(* IEC 61131-3 sources: canworks/examples/virtual-plant/pous/programs, 3 files *)

(* ---- canworks_in.st ---- *)
PROGRAM canworks_in
  VAR
    i0  : WORD AT %IW100; (* cw_map_hash *)
    i1  : WORD AT %IW101; (* cw_map_hash_w1 *)
    i2  : WORD AT %IW102; (* cw_status *)
    i3  : WORD AT %IW103; (* cw_status_w1 *)
    i4  : WORD AT %IW104; (* cw_status_w2 *)
    i5  : WORD AT %IW105; (* cw_status_w3 *)
    i6  : WORD AT %IW106; (* io_rtd_AI0_Input_PV *)
    i7  : WORD AT %IW107; (* io_rtd_AI1_Input_PV *)
    i8  : WORD AT %IW108; (* io_rtd_AI2_Input_PV *)
    i9  : WORD AT %IW109; (* io_rtd_AI3_Input_PV *)
    i10 : WORD AT %IW110; (* io_dio_Read_input_8_bit_1 *)
    i11 : WORD AT %IW111; (* io_dio_Read_analogue_input_1 *)
    i12 : WORD AT %IW112; (* io_dio_Read_analogue_input_2 *)
    i13 : WORD AT %IW113; (* io_dio_operating_hours *)
    i14 : WORD AT %IW114; (* io_dio_operating_hours_w1 *)
    i15 : WORD AT %IW115; (* io_new_io_Read_input_8_bit_1 *)
    i16 : WORD AT %IW116; (* motion_conveyor_speed_actual *)
    i17 : WORD AT %IW117; (* motion_conveyor_belt_position *)
    i18 : WORD AT %IW118; (* motion_conveyor_belt_position_w1 *)
    i19 : WORD AT %IW119; (* host_cell_alarm *)
    i20 : WORD AT %IW120; (* cell_temp_limit *)
    i21 : WORD AT %IW121; (* host_cell_belt_position *)
    i22 : WORD AT %IW122; (* host_cell_belt_position_w1 *)
    i23 : WORD AT %IW123; (* host_cell_cycle_count *)
    i24 : WORD AT %IW124; (* host_cell_cycle_count_w1 *)
    i25 : WORD AT %IW125; (* host_cell_temperature *)
    i26 : WORD AT %IW126; (* host_cell_Nodes_0_31 *)
    i27 : WORD AT %IW127; (* host_cell_Nodes_0_31_w1 *)
    i28 : WORD AT %IW128; (* host_cell_Nodes_0_31_2 *)
    i29 : WORD AT %IW129; (* host_cell_Nodes_0_31_2_w1 *)
    i30 : WORD AT %IW130; (* io_can_bus_state *)
    i31 : WORD AT %IW131; (* io_rtd_ok *)
    i32 : WORD AT %IW132; (* io_rtd_emcy *)
    i33 : WORD AT %IW133; (* io_dio_state *)
    i34 : WORD AT %IW134; (* io_dio_emcy *)
    i35 : WORD AT %IW135; (* io_dio_operating_hours_status *)
    i36 : WORD AT %IW136; (* motion_can_master_state *)
    i37 : WORD AT %IW137; (* motion_conveyor_emcy *)
    i38 : WORD AT %IW138; (* host_can_master_state *)
    i39 : WORD AT %IW139; (* host_cell_state *)
    i40 : WORD AT %IW140; (* host_cell_emcy *)
    i41 : WORD AT %IW141; (* cw_live_list_io *)
    i42 : WORD AT %IW142; (* cw_live_list_io_w1 *)
    i43 : WORD AT %IW143; (* cw_live_list_io_w2 *)
    i44 : WORD AT %IW144; (* cw_live_list_io_w3 *)
    i45 : WORD AT %IW145; (* cw_live_list_io_w4 *)
    i46 : WORD AT %IW146; (* cw_live_list_io_w5 *)
    i47 : WORD AT %IW147; (* cw_live_list_io_w6 *)
    i48 : WORD AT %IW148; (* cw_live_list_io_w7 *)
    i49 : WORD AT %IW149; (* cw_live_list_motion *)
    i50 : WORD AT %IW150; (* cw_live_list_motion_w1 *)
    i51 : WORD AT %IW151; (* cw_live_list_motion_w2 *)
    i52 : WORD AT %IW152; (* cw_live_list_motion_w3 *)
    i53 : WORD AT %IW153; (* cw_live_list_motion_w4 *)
    i54 : WORD AT %IW154; (* cw_live_list_motion_w5 *)
    i55 : WORD AT %IW155; (* cw_live_list_motion_w6 *)
    i56 : WORD AT %IW156; (* cw_live_list_motion_w7 *)
    i57 : WORD AT %IW157; (* cw_live_list_host *)
    i58 : WORD AT %IW158; (* cw_live_list_host_w1 *)
    i59 : WORD AT %IW159; (* cw_live_list_host_w2 *)
    i60 : WORD AT %IW160; (* cw_live_list_host_w3 *)
    i61 : WORD AT %IW161; (* cw_live_list_host_w4 *)
    i62 : WORD AT %IW162; (* cw_live_list_host_w5 *)
    i63 : WORD AT %IW163; (* cw_live_list_host_w6 *)
    i64 : WORD AT %IW164; (* cw_live_list_host_w7 *)
    i65 : WORD AT %IW165; (* cw_sdo_bridge_response *)
    i66 : WORD AT %IW166; (* cw_sdo_bridge_response_w1 *)
    i67 : WORD AT %IW167; (* cw_sdo_bridge_response_w2 *)
    i68 : WORD AT %IW168; (* cw_sdo_bridge_response_w3 *)
    i69 : WORD AT %IW169; (* cw_sdo_bridge_response_w4 *)
    i70 : WORD AT %IW170; (* cw_sdo_bridge_response_w5 *)
    i71 : WORD AT %IW171; (* cw_sdo_bridge_response_w6 *)
  END_VAR
  VAR
    last_counter : WORD;
    moved        : BOOL;
    stale        : TON;
  END_VAR

(* Generated by canworks from canworks/canworks.json: do not edit, Save rewrites it. *)
moved := i3 <> last_counter;
last_counter := i3;
stale(IN := NOT moved, PT := T#300ms);
canworks.ok := i0 = WORD#16#662D AND i1 = WORD#16#449C AND NOT stale.Q;
canworks.bus_ok := canworks.ok AND (i5 AND WORD#16#0002) = WORD#0;
canworks.link[21] := WORD#16#0B06 OR SEL(canworks.ok, WORD#0, WORD#1);
canworks.link[0] := i2;
canworks.link[1] := i3;
canworks.link[2] := i4;
canworks.link[3] := i5;
canworks.link[14] := i65;
canworks.link[15] := i66;
canworks.link[16] := i67;
canworks.link[17] := i68;
canworks.link[18] := i69;
canworks.link[19] := i70;
canworks.link[20] := i71;
canworks.link[25] := i41;
canworks.link[26] := i42;
canworks.link[27] := i43;
canworks.link[28] := i44;
canworks.link[29] := i45;
canworks.link[30] := i46;
canworks.link[31] := i47;
canworks.link[32] := i48;
canworks.link[33] := i49;
canworks.link[34] := i50;
canworks.link[35] := i51;
canworks.link[36] := i52;
canworks.link[37] := i53;
canworks.link[38] := i54;
canworks.link[39] := i55;
canworks.link[40] := i56;
canworks.link[49] := i57;
canworks.link[50] := i58;
canworks.link[51] := i59;
canworks.link[52] := i60;
canworks.link[53] := i61;
canworks.link[54] := i62;
canworks.link[55] := i63;
canworks.link[56] := i64;
canworks.io_can_bus_state := SEL(canworks.ok, USINT#0, WORD_TO_USINT((i30 AND WORD#16#00FF)));
canworks.io_can_master_state := SEL(canworks.ok, USINT#0, WORD_TO_USINT(SHR(i30, 8)));
canworks.motion_can_master_state := SEL(canworks.ok, USINT#0, WORD_TO_USINT(SHR(i36, 8)));
canworks.host_can_master_state := SEL(canworks.ok, USINT#0, WORD_TO_USINT((i38 AND WORD#16#00FF)));
canworks.io_rtd_ok := SEL(canworks.ok, FALSE, (i31 AND WORD#16#0100) <> WORD#0);
canworks.io_rtd_state := SEL(canworks.ok, USINT#0, WORD_TO_USINT((i31 AND WORD#16#00FF)));
canworks.io_rtd_emcy := SEL(canworks.ok, WORD#0, i32);
canworks.io_rtd_tpdo1_timeout := SEL(canworks.ok, FALSE, (i31 AND WORD#16#0200) <> WORD#0);
canworks.io_rtd_AI0_Input_PV := WORD_TO_INT(i6);
canworks.io_rtd_AI1_Input_PV := WORD_TO_INT(i7);
canworks.io_rtd_AI2_Input_PV := WORD_TO_INT(i8);
canworks.io_rtd_AI3_Input_PV := WORD_TO_INT(i9);
canworks.io_dio_ok := SEL(canworks.ok, FALSE, (i31 AND WORD#16#0400) <> WORD#0);
canworks.io_dio_state := SEL(canworks.ok, USINT#0, WORD_TO_USINT(SHR(i33, 8)));
canworks.io_dio_emcy := SEL(canworks.ok, WORD#0, i34);
canworks.io_dio_Read_input_8_bit_1 := WORD_TO_USINT(SHR(i10, 8));
canworks.io_dio_Read_input_8_bit_2 := WORD_TO_USINT((i10 AND WORD#16#00FF));
canworks.io_dio_Read_analogue_input_1 := WORD_TO_INT(i11);
canworks.io_dio_Read_analogue_input_2 := WORD_TO_INT(i12);
canworks.io_dio_operating_hours := DWORD_TO_UDINT((SHL(WORD_TO_DWORD(i14), 16) OR WORD_TO_DWORD(i13)));
canworks.io_dio_operating_hours_status := SEL(canworks.ok, USINT#0, WORD_TO_USINT(SHR(i35, 8)));
canworks.io_dio_filter_time_status := SEL(canworks.ok, USINT#0, WORD_TO_USINT((i35 AND WORD#16#00FF)));
canworks.io_new_io_ok := SEL(canworks.ok, FALSE, (i31 AND WORD#16#0800) <> WORD#0);
canworks.io_new_io_Read_input_8_bit_1 := WORD_TO_USINT(SHR(i15, 8));
canworks.motion_conveyor_ok := SEL(canworks.ok, FALSE, (i31 AND WORD#16#1000) <> WORD#0);
canworks.motion_conveyor_state := SEL(canworks.ok, USINT#0, WORD_TO_USINT((i36 AND WORD#16#00FF)));
canworks.motion_conveyor_emcy := SEL(canworks.ok, WORD#0, i37);
canworks.motion_conveyor_speed_actual := WORD_TO_INT(i16);
canworks.motion_conveyor_belt_position := DWORD_TO_DINT((SHL(WORD_TO_DWORD(i18), 16) OR WORD_TO_DWORD(i17)));
canworks.host_cell_ok := SEL(canworks.ok, FALSE, (i31 AND WORD#16#4000) <> WORD#0);
canworks.host_cell_state := SEL(canworks.ok, USINT#0, WORD_TO_USINT(SHR(i39, 8)));
canworks.host_cell_emcy := SEL(canworks.ok, WORD#0, i40);
canworks.host_cell_alarm := (i19 AND WORD#16#0200) <> WORD#0;
canworks.host_cell_belt_position := DWORD_TO_DINT((SHL(WORD_TO_DWORD(i22), 16) OR WORD_TO_DWORD(i21)));
canworks.host_cell_cycle_count := DWORD_TO_UDINT((SHL(WORD_TO_DWORD(i24), 16) OR WORD_TO_DWORD(i23)));
canworks.host_cell_temperature := WORD_TO_INT(i25);
canworks.host_cell_Nodes_0_31 := DWORD_TO_UDINT((SHL(WORD_TO_DWORD(i27), 16) OR WORD_TO_DWORD(i26)));
canworks.host_cell_Nodes_0_31_2 := DWORD_TO_UDINT((SHL(WORD_TO_DWORD(i29), 16) OR WORD_TO_DWORD(i28)));
canworks.cell_line_run := (i19 AND WORD#16#0100) <> WORD#0;
canworks.cell_temp_limit := WORD_TO_INT(i20);
canworks.cell_state := SEL(canworks.ok, USINT#0, WORD_TO_USINT(SHR(i38, 8)));
canworks.cell_comm_ok := SEL(canworks.ok, FALSE, (i31 AND WORD#16#2000) <> WORD#0);

END_PROGRAM

(* ---- canworks_out.st ---- *)
PROGRAM canworks_out
  VAR
    q0  : WORD AT %QW100; (* cw_plc_link *)
    q1  : WORD AT %QW101; (* cw_plc_link_w1 *)
    q2  : WORD AT %QW102; (* cw_plc_link_w2 *)
    q3  : WORD AT %QW103; (* io_dio_Write_output_8_bit_1 *)
    q4  : WORD AT %QW104; (* io_dio_Write_analogue_output_2 *)
    q5  : WORD AT %QW105; (* io_dio_filter_time *)
    q6  : WORD AT %QW106; (* io_new_io_Write_output_8_bit_1 *)
    q7  : WORD AT %QW107; (* motion_conveyor_speed_setpoint *)
    q8  : WORD AT %QW108; (* host_cell_line_run *)
    q9  : WORD AT %QW109; (* cell_belt_position *)
    q10 : WORD AT %QW110; (* cell_belt_position_w1 *)
    q11 : WORD AT %QW111; (* cell_cycle_count *)
    q12 : WORD AT %QW112; (* cell_cycle_count_w1 *)
    q13 : WORD AT %QW113; (* host_cell_temp_limit *)
    q14 : WORD AT %QW114; (* host_cell_analog_out *)
    q15 : WORD AT %QW115; (* io_dio_filter_time_trig *)
    q16 : WORD AT %QW116; (* cell_emcy *)
    q17 : WORD AT %QW117; (* cell_errreg *)
    q18 : WORD AT %QW118; (* cw_control *)
    q19 : WORD AT %QW119; (* cw_control_w1 *)
    q20 : WORD AT %QW120; (* cw_control_w2 *)
    q21 : WORD AT %QW121; (* cw_sdo_bridge_request *)
    q22 : WORD AT %QW122; (* cw_sdo_bridge_request_w1 *)
    q23 : WORD AT %QW123; (* cw_sdo_bridge_request_w2 *)
    q24 : WORD AT %QW124; (* cw_sdo_bridge_request_w3 *)
    q25 : WORD AT %QW125; (* cw_sdo_bridge_request_w4 *)
    q26 : WORD AT %QW126; (* cw_sdo_bridge_request_w5 *)
    q27 : WORD AT %QW127; (* cw_sdo_bridge_request_w6 *)
  END_VAR
  VAR
    d9  : DWORD;
    d11 : DWORD;
  END_VAR

(* Generated by canworks from canworks/canworks.json: do not edit, Save rewrites it. *)
d9 := DINT_TO_DWORD(canworks.cell_belt_position);
d11 := UDINT_TO_DWORD(canworks.cell_cycle_count);
q3 := SHL((USINT_TO_WORD(canworks.io_dio_Write_output_8_bit_1) AND WORD#16#00FF), 8) OR (USINT_TO_WORD(canworks.io_dio_Write_output_8_bit_2) AND WORD#16#00FF);
q4 := INT_TO_WORD(canworks.io_dio_Write_analogue_output_2);
q5 := UINT_TO_WORD(canworks.io_dio_filter_time);
q6 := SHL((USINT_TO_WORD(canworks.io_new_io_Write_output_8_bit_1) AND WORD#16#00FF), 8);
q7 := INT_TO_WORD(canworks.motion_conveyor_speed_setpoint);
q8 := SEL(canworks.host_cell_line_run, WORD#0, WORD#16#0200) OR SEL(canworks.cell_alarm, WORD#0, WORD#16#0100);
q9 := DWORD_TO_WORD(d9);
q10 := DWORD_TO_WORD(SHR(d9, 16));
q11 := DWORD_TO_WORD(d11);
q12 := DWORD_TO_WORD(SHR(d11, 16));
q13 := INT_TO_WORD(canworks.host_cell_temp_limit);
q14 := INT_TO_WORD(canworks.host_cell_analog_out);
q15 := SEL(canworks.io_dio_filter_time_trig, WORD#0, WORD#16#0100);
q16 := canworks.cell_emcy;
q17 := SHL((BYTE_TO_WORD(canworks.cell_errreg) AND WORD#16#00FF), 8);
q18 := canworks.link[4];
q19 := canworks.link[5];
q20 := canworks.link[6];
q21 := canworks.link[7];
q22 := canworks.link[8];
q23 := canworks.link[9];
q24 := canworks.link[10];
q25 := canworks.link[11];
q26 := canworks.link[12];
q27 := canworks.link[13];
(* PLC link header, last: running, then the map hash 0x662d449c *)
q1 := WORD#16#662D;
q2 := WORD#16#449C;
q0 := WORD#1;

END_PROGRAM

(* ---- main.st ---- *)
PROGRAM main
  VAR
    (* The demo (docs/tour.md). The CANopen values are in the `canworks`
       variable list, which canworks_in fills from the bridge before main and
       canworks_out sends after it (the configurator writes all three). *)
    temp_c          : REAL;   (* RTD channel 0 in degC (the module sends 0.1 degC) *)
    limit           : INT;    (* alarm limit in 0.1 degC, from the cell's upper master *)
    alarm           : BOOL;   (* channel 0 above the limit: DIO-16 output 0.0 and the cell's alarm *)
    fault           : BOOL;   (* a node lost, a PDO timed out or an EMCY active: new_io output 0.0 *)
    pattern         : USINT := 1;  (* running light on DIO-16 output byte 2, read back on input byte 2 *)
    tick            : INT;
    loop_errors     : UDINT;  (* times the read-back input did not follow the output *)
    loop_ok         : BOOL;
    cycles          : UDINT;
    restart_dio     : BOOL;   (* set it in the debugger: NMT reset of node dio (6) *)
    started         : BOOL;
    rd_product      : CO_SDO_READ;   (* network io (0), node 5: 0x1018:2 product code *)
    rd_conveyor     : CO_SDO_READ;   (* network motion (1), node 4: 0x1018:2 product code *)
    wr_ai_interrupt : CO_SDO_WRITE;  (* network io (0), node 6: 0x6423 analogue input global interrupt enable *)
    reset_dio       : CO_NMT;        (* network io (0), node 6: RESET NODE when restart_dio is set *)
    rtd_product     : UDINT;
    conveyor_product : UDINT;
    sdo_errors      : INT;
    (* The host network plays the cell's machine controller (the upper master). *)
    host_field_ok   : BOOL;   (* the gateway reports io nodes 5, 6, 7 and motion node 4 operational *)
    speed           : INT := 1000;  (* conveyor speed while the upper master runs the line *)
  END_VAR

(* Temperature, alarm and the I/O loopback on network io *)
cycles := cycles + 1;
canworks.cell_cycle_count := cycles;
temp_c := INT_TO_REAL(canworks.io_rtd_AI0_Input_PV) / 10.0;
limit := canworks.cell_temp_limit;
IF limit = 0 THEN limit := 250; END_IF  (* no upper master: 25.0 degC *)
alarm := canworks.io_rtd_ok AND canworks.io_rtd_AI0_Input_PV > limit;
canworks.cell_alarm := alarm;
IF alarm THEN
  canworks.cell_emcy := 16#4210;  (* temperature too high: the cell slave sends it once *)
  canworks.cell_errreg := 16#09;  (* generic + temperature *)
ELSE
  canworks.cell_emcy := 0;
  canworks.cell_errreg := 0;
END_IF
canworks.io_dio_Write_output_8_bit_1 := BOOL_TO_USINT(alarm);

(* DIO-16 loops its outputs back to its inputs: a running light on byte 2,
   checked a few PDO round trips later. *)
tick := tick + 1;
IF tick >= 25 THEN
  tick := 0;
  IF canworks.io_dio_ok THEN
    loop_ok := canworks.io_dio_Read_input_8_bit_2 = pattern;
    IF NOT loop_ok THEN loop_errors := loop_errors + 1; END_IF
  END_IF
  pattern := ROL(pattern, 1);
END_IF
canworks.io_dio_Write_output_8_bit_2 := pattern;
canworks.io_dio_Write_analogue_output_2 := canworks.io_rtd_AI1_Input_PV;  (* AO 2 follows RTD channel 1 *)

(* Reactions: lost nodes, the RTD PDO's receive timeout, EMCYs *)
fault := NOT canworks.io_rtd_ok OR NOT canworks.io_dio_ok OR NOT canworks.motion_conveyor_ok
         OR canworks.io_rtd_tpdo1_timeout
         OR canworks.io_rtd_emcy <> 0 OR canworks.io_dio_emcy <> 0 OR canworks.motion_conveyor_emcy <> 0;
canworks.io_new_io_Write_output_8_bit_1 := BOOL_TO_USINT(fault) OR SHL(BOOL_TO_USINT(NOT host_field_ok), 1);

(* NMT: restart_dio resets node 6 once (set it again for another reset). *)
reset_dio(EXECUTE := restart_dio, NETWORK := 0, NODE := 6, COMMAND := 129, LINK := canworks.link);
IF reset_dio.DONE OR reset_dio.ERROR THEN restart_dio := FALSE; END_IF

(* SDO: read and write once after the nodes are up (again after a node comes
   back). *)
started := canworks.ok AND canworks.io_rtd_ok AND canworks.io_dio_ok AND canworks.motion_conveyor_ok;
rd_product(EXECUTE := started, NETWORK := 0, NODE := 5, INDEX := 16#1018, SUBINDEX := 2, LINK := canworks.link);
IF rd_product.DONE THEN rtd_product := rd_product.DATA; END_IF
rd_conveyor(EXECUTE := started, NETWORK := 1, NODE := 4, INDEX := 16#1018, SUBINDEX := 2, LINK := canworks.link);
IF rd_conveyor.DONE THEN conveyor_product := rd_conveyor.DATA; END_IF
wr_ai_interrupt(EXECUTE := started, NETWORK := 0, NODE := 6, INDEX := 16#6423, SUBINDEX := 0,
                DATA := 1, SIZE := 1, LINK := canworks.link);
IF rd_product.ERROR OR rd_conveyor.ERROR OR wr_ai_interrupt.ERROR THEN sdo_errors := sdo_errors + 1; END_IF

(* The host network: the cell's machine controller. It runs the line, sets
   the alarm limit and sends the temperature it gets through the gateway
   back down to DIO-16's analogue output 1. *)
canworks.host_cell_line_run := canworks.host_cell_ok;
canworks.host_cell_temp_limit := 250;
canworks.host_cell_analog_out := canworks.host_cell_temperature;
host_field_ok := canworks.host_cell_ok AND (canworks.host_cell_Nodes_0_31 AND 16#E0) = 16#E0
                 AND (canworks.host_cell_Nodes_0_31_2 AND 16#10) = 16#10;

(* The conveyor runs while the upper master runs the line; its belt position
   goes up to the host. *)
IF canworks.cell_line_run AND canworks.motion_conveyor_ok THEN
  canworks.motion_conveyor_speed_setpoint := speed;
ELSE
  canworks.motion_conveyor_speed_setpoint := 0;
END_IF
canworks.cell_belt_position := canworks.motion_conveyor_belt_position;

END_PROGRAM
